// TIA Portal V20 export
Screen "PopupCycleTimeLegend"  360x155
  ScreenItem "Textfeld_Legende" at 61,2 size 209x25  Type=HmiTextBox
  ScreenItem "Textfeld_3" at 10,37 size 140x20  Type=HmiTextBox
  ScreenItem "Textfeld_11" at 155,37 size 145x20  Type=HmiTextBox
  ScreenItem "Cancel Mode" at 288,1 size 71x42  Type=HmiButton
  ScreenItem "Textfeld_5" at 0,0 size 140x20  Type=HmiTextBox
  ScreenItem "Textfeld_13" at 145,1 size 200x20  Type=HmiTextBox
  ScreenItem "Textfeld_4" at 0,0 size 140x20  Type=HmiTextBox
  ScreenItem "Textfeld_12" at 145,1 size 202x20  Type=HmiTextBox
  ScreenItem "Textfeld_6" at 0,0 size 140x20  Type=HmiTextBox
  ScreenItem "Textfeld_14" at 145,1 size 200x20  Type=HmiTextBox
  ScreenItem "Textfeld_1" at 0,0 size 140x20  Type=HmiTextBox
  ScreenItem "Textfeld_9" at 145,1 size 200x20  Type=HmiTextBox
